FUNCTION_BLOCK Q_StringValue (* Command Change String Value ( Part 6 - F.24 ) *)
  (* Standard: ISO 11783-6; Description: This command sends a string to the VT. The length of the string including '\0' may not be longer than the define ISO_VTC_CMD_STR_MAX_LENGTH. Take care that '\0' is trailed. Return values iso_s16 - E_NO_ERR ( 0 )  - transport started - E_OVERFLOW (-6 ) - buffer overflow - E_NOACT (-8 ) - Command not possible in current state - E_NO_INSTANCE (-21) - No VT client available *)
  (* Version 1.0, 2022-07-08, franz *)
  (* Documentation:
  This command sends a string to the VT. The length of the string including '' may not be longer than the define ISO_VTC_CMD_STR_MAX_LENGTH. Take care that '' is trailed.
   Return values
   iso_s16
    - E_NO_ERR ( 0 )  - transport started
   - E_OVERFLOW (-6 ) - buffer overflow
   - E_NOACT (-8 ) - Command not possible in current state
   - E_NO_INSTANCE (-21) - No VT client available
  *)
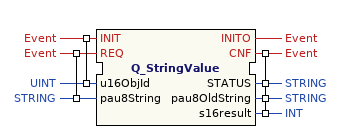
  EVENT_INPUT
    INIT WITH u16ObjId; (* Service Initialization *)
    REQ WITH pau8String; (* Service Request *)
  END_EVENT
  EVENT_OUTPUT
    INITO; (* Initialization Confirm *)
    CNF WITH STATUS, pau8OldString, s16result; (* Confirmation of Requested Service *)
  END_EVENT
  VAR_INPUT
    u16ObjId : UINT; (* Object ID *)
    pau8String : STRING; (* Pointer to string *)
  END_VAR
  VAR_OUTPUT
    STATUS : STRING; (* Service Status *)
    pau8OldString : STRING; (* Old pointer to string *)
    s16result : INT; (* retval see description *)
  END_VAR
END_FUNCTION_BLOCK
